FUNCTION "FRK_UnitRelease" : Void
{ S7_Optimized_Access := 'TRUE' }
VERSION : 0.1
VAR_INPUT
    Gate : DInt;
    Desired : DInt;
    Trusted : Bool;
    Core : "FRK_Core";
    Unit : "FRK_Unit";
    Status : "ST_ModuleStatus";
    Policy : Array[0..6] of "ST_ModePolicy";
    Access : "FRK_Access";
    Supported : Array[0..6] of Bool;
END_VAR
VAR_IN_OUT
    Report : "ST_ReleaseReport";
END_VAR
BEGIN
    #Report.Count := 0;
    #Report.Released := TRUE;
    IF #Gate <> 5 AND #Gate <> 4
        AND #Gate <> 7 AND #Gate <> 2
        AND #Gate <> 8
        AND NOT (#Unit.ConfigEnabled AND #Gate = 1)
        AND NOT (#Unit.ConfigSetsEnabled AND #Gate = 11)
        AND NOT (#Unit.ModelEnabled AND #Gate = 3) THEN
        "FRK_ReleaseReason"(Report := #Report, Description := WSTRING#'std.error.unsupportedHmiRequest', Reason := 2008, Path := STRING_TO_WSTRING(#Status.Name), Kind := 4);
        RETURN;
    END_IF;
    IF NOT #Trusted THEN
        IF #Access.CurrentLevel < #Access.Policy.Required[#Gate] THEN
            "FRK_ReleaseReason"(Report := #Report, Description := WSTRING#'std.release.insufficientAction', Reason := 2002, Path := STRING_TO_WSTRING(#Status.Name), Kind := 1);
        END_IF;
    END_IF;
    CASE #Gate OF
        3:
            IF #Core.Exec <> 0 OR #Unit.ModePending OR #Unit.Clearing OR NOT "FRK_DescendantsReady"(OwnerIndex := #Core.RegIndex) THEN
                "FRK_ReleaseReason"(Report := #Report, Description := WSTRING#'std.error.hmiRequestRejected', Reason := 2011, Path := STRING_TO_WSTRING(#Status.Name), Kind := 4);
            END_IF;
            IF #Unit.AlarmBlocking THEN
                "FRK_ReleaseReason"(Report := #Report, Description := WSTRING#'std.release.manualReset', Reason := 0, Path := STRING_TO_WSTRING(#Status.Name), Kind := 2);
            END_IF;
            IF NOT #Unit.Permit THEN
                "FRK_ReleaseReason"(Report := #Report, Description := #Unit.PermitDiag.Description, Reason := #Unit.PermitDiag.ReasonCode, Path := #Unit.PermitDiag.SourcePath, Kind := 3);
            END_IF;
        5:
            // Desired=0 is Start, Desired=1 is Stop. Generic action query is Stop.
            IF #Desired = 0 THEN
                IF #Unit.Mode = 1 OR #Unit.ModePending THEN
                    "FRK_ReleaseReason"(Report := #Report, Description := WSTRING#'std.error.unsupportedModeRequest', Reason := 2002, Path := STRING_TO_WSTRING(#Status.Name), Kind := 0);
                END_IF;
                IF #Core.Exec <> 0 OR #Unit.RunReq OR #Unit.Clearing OR #Unit.FaultLatched THEN
                    "FRK_ReleaseReason"(Report := #Report, Description := WSTRING#'std.error.hmiRequestRejected', Reason := 2011, Path := STRING_TO_WSTRING(#Status.Name), Kind := 4);
                END_IF;
                IF #Unit.AlarmBlocking THEN
                    "FRK_ReleaseReason"(Report := #Report, Description := WSTRING#'std.release.manualReset', Reason := 0, Path := STRING_TO_WSTRING(#Status.Name), Kind := 2);
                END_IF;
                IF #Unit.ConfigBlocked THEN
                    "FRK_ReleaseReason"(Report := #Report, Description := WSTRING#'std.release.configRestoreUnacknowledged', Reason := 2040, Path := STRING_TO_WSTRING(#Status.Name), Kind := 2);
                END_IF;
                IF NOT #Unit.Permit THEN
                    "FRK_ReleaseReason"(Report := #Report, Description := #Unit.PermitDiag.Description, Reason := #Unit.PermitDiag.ReasonCode, Path := #Unit.PermitDiag.SourcePath, Kind := 3);
                END_IF;
            END_IF;
        4:
            IF #Unit.ModePending THEN
                "FRK_ReleaseReason"(Report := #Report, Description := WSTRING#'std.release.modeChangeAlreadyPending', Reason := 2011, Path := STRING_TO_WSTRING(#Status.Name), Kind := 0);
            END_IF;
            IF #Core.Exec = 1 AND #Unit.Mode <> 1 THEN
                IF #Policy[#Unit.Mode].Shield = 2 THEN
                    "FRK_ReleaseReason"(Report := #Report, Description := WSTRING#'std.release.modeSwitchBlockedWhileRunning', Reason := 2002, Path := STRING_TO_WSTRING(#Status.Name), Kind := 0);
                END_IF;
            END_IF;
            IF #Desired <> -1 THEN
                IF #Desired < 0 OR #Desired >= 7 THEN
                    "FRK_ReleaseReason"(Report := #Report, Description := WSTRING#'std.error.unsupportedModeRequest', Reason := 2008, Path := STRING_TO_WSTRING(#Status.Name), Kind := 0);
                ELSIF NOT #Supported[#Desired] THEN
                    "FRK_ReleaseReason"(Report := #Report, Description := WSTRING#'std.error.unsupportedModeRequest', Reason := 2008, Path := STRING_TO_WSTRING(#Status.Name), Kind := 0);
                END_IF;
            END_IF;
        7:
            // The complete alarm model is separate; this gate owns the current latch.
            IF NOT #Unit.FaultLatched AND NOT #Unit.AlarmBlocking AND #Core.Exec = 0 AND NOT #Unit.Clearing AND NOT #Unit.ModePending AND NOT #Unit.FollowStart THEN
                IF "FRK_DescendantsReady"(OwnerIndex := #Core.RegIndex) THEN
                    "FRK_ReleaseReason"(Report := #Report, Description := WSTRING#'std.release.noBlockingAlarm', Reason := 2011, Path := STRING_TO_WSTRING(#Status.Name), Kind := 4);
                END_IF;
            END_IF;
        2:
            "FRK_ManualCommon"(Core := #Core, Unit := #Unit, Status := #Status, Report := #Report);
        ELSE
            RETURN;
    END_CASE;
END_FUNCTION

FUNCTION "FRK_ManualCommon" : Void
{ S7_Optimized_Access := 'TRUE' }
VERSION : 0.1
VAR_INPUT
    Core : "FRK_Core";
    Unit : "FRK_Unit";
    Status : "ST_ModuleStatus";
END_VAR
VAR_IN_OUT
    Report : "ST_ReleaseReport";
END_VAR
BEGIN
    IF #Unit.Mode <> 1 OR #Unit.ModePending THEN
        "FRK_ReleaseReason"(Report := #Report, Description := WSTRING#'std.release.manualModeRequired', Reason := 2002, Path := STRING_TO_WSTRING(#Status.Name), Kind := 0);
    END_IF;
    IF #Core.Exec <> 0 OR #Unit.Clearing OR #Unit.FaultLatched THEN
        "FRK_ReleaseReason"(Report := #Report, Description := WSTRING#'std.error.hmiRequestRejected', Reason := 2011, Path := STRING_TO_WSTRING(#Status.Name), Kind := 4);
    END_IF;
    IF #Unit.AlarmBlocking THEN
        "FRK_ReleaseReason"(Report := #Report, Description := WSTRING#'std.release.manualReset', Reason := 0, Path := STRING_TO_WSTRING(#Status.Name), Kind := 2);
    END_IF;
    IF NOT #Unit.Permit THEN
        "FRK_ReleaseReason"(Report := #Report, Description := #Unit.PermitDiag.Description, Reason := #Unit.PermitDiag.ReasonCode, Path := #Unit.PermitDiag.SourcePath, Kind := 3);
    END_IF;
END_FUNCTION

FUNCTION "FRK_ManualCondition" : Void
{ S7_Optimized_Access := 'TRUE' }
VERSION : 0.1
VAR_INPUT
    Slot : Int;
    Value : DInt;
    Ok : Bool;
    Diag : "ST_Diagnostic";
    Bypassable : Bool;
END_VAR
VAR_IN_OUT
    Conditions : Array[1..16] of "FRK_ManualConditionRow";
END_VAR
BEGIN
    IF #Slot < 1 OR #Slot > 16 THEN RETURN; END_IF;
    #Conditions[#Slot].Used := TRUE;
    #Conditions[#Slot].Value := #Value;
    #Conditions[#Slot].Ok := #Ok;
    #Conditions[#Slot].Diag := #Diag;
    #Conditions[#Slot].Bypassable := #Bypassable;
END_FUNCTION

FUNCTION "FRK_ManualApply" : Void
{ S7_Optimized_Access := 'TRUE' }
VERSION : 0.1
VAR_INPUT
    Request : "ST_HmiRequest";
    Status : "ST_ModuleStatus";
    Core : "FRK_Core";
    Commands : Array[1..12] of "ST_CommandInfo";
    Count : DInt;
    Conditions : Array[1..16] of "FRK_ManualConditionRow";
END_VAR
VAR_IN_OUT
    Report : "ST_ReleaseReport";
    Execute : Bool;
    Command : DInt;
    ManualOwned : Bool;
END_VAR
VAR_TEMP
    Index : Int;
    Supported : Bool;
    PreviousCount : Int;
END_VAR
BEGIN
    #Supported := FALSE;
    IF #Count >= 0 AND #Count <= 12 THEN
        FOR #Index := 1 TO DINT_TO_INT(#Count) DO
            IF #Commands[#Index].Value = #Request.IntValue AND #Commands[#Index].Style = 0 THEN #Supported := TRUE; END_IF;
        END_FOR;
    END_IF;
    IF NOT #Supported THEN
        "FRK_ReleaseReason"(Report := #Report, Description := WSTRING#'std.error.unsupportedHmiRequest', Reason := 2008, Path := STRING_TO_WSTRING(#Status.Name), Kind := 4);
    END_IF;
    IF #Core.Exec <> 0 OR #Execute OR #Core.ReleasePending THEN
        "FRK_ReleaseReason"(Report := #Report, Description := WSTRING#'std.error.hmiRequestRejected', Reason := 2011, Path := STRING_TO_WSTRING(#Status.Name), Kind := 4);
    END_IF;
    FOR #Index := 1 TO 16 DO
        IF #Conditions[#Index].Used AND NOT #Conditions[#Index].Ok THEN
            IF #Conditions[#Index].Value = 0 OR #Conditions[#Index].Value = #Request.IntValue THEN
                #PreviousCount := #Report.Count;
                "FRK_ReleaseReason"(Report := #Report, Description := #Conditions[#Index].Diag.Description, Reason := #Conditions[#Index].Diag.ReasonCode, Path := STRING_TO_WSTRING(#Status.Name), Kind := 3);
                IF #Report.Count > #PreviousCount THEN #Report.Reasons[#Report.Count].Bypassable := #Conditions[#Index].Bypassable; END_IF;
            END_IF;
        END_IF;
    END_FOR;
    IF #Request.Kind = 11 AND #Report.Released THEN
        #Command := #Request.IntValue;
        #Execute := TRUE;
        #ManualOwned := TRUE;
    END_IF;
END_FUNCTION

FUNCTION "FRK_ManualFinish" : Void
{ S7_Optimized_Access := 'TRUE' }
VERSION : 0.1
VAR_INPUT
    Core : "FRK_Core";
END_VAR
VAR_IN_OUT
    Execute : Bool;
    ManualOwned : Bool;
END_VAR
BEGIN
    IF #ManualOwned AND #Core.Exec <> 1 THEN
        #Execute := FALSE;
        #ManualOwned := FALSE;
    END_IF;
END_FUNCTION

FUNCTION "FRK_UnitCascade" : Void
{ S7_Optimized_Access := 'TRUE' }
VERSION : 0.1
VAR_INPUT
    ParentUnit : "FRK_Unit";
    Supported : Array[0..6] of Bool;
END_VAR
VAR_IN_OUT
    Core : "FRK_Core";
    Unit : "FRK_Unit";
    Status : "ST_ModuleStatus";
    Policy : Array[0..6] of "ST_ModePolicy";
    Access : "FRK_Access";
    AlarmLog : "FRK_AlarmLog";
END_VAR
VAR_TEMP
    Request : "ST_HmiRequest";
END_VAR
BEGIN
    IF NOT #ParentUnit.CascadePending THEN RETURN; END_IF;
    IF #ParentUnit.CascadeKind = 6 OR #ParentUnit.CascadeKind = 9 THEN
        #Unit.FollowStart := FALSE;
        #Request.Kind := #ParentUnit.CascadeKind;
        "FRK_UnitOperation"(Core := #Core, Unit := #Unit, Status := #Status, Policy := #Policy, Access := #Access, Supported := #Supported, Request := #Request, Response := "FRK_UnitScratch".Response, Trusted := TRUE);
        RETURN;
    END_IF;
    #Request.Kind := 3;
    #Request.IntValue := #ParentUnit.CascadeMode;
    "FRK_UnitOperation"(Core := #Core, Unit := #Unit, Status := #Status, Policy := #Policy, Access := #Access, Supported := #Supported, Request := #Request, Response := "FRK_UnitScratch".Response, Trusted := TRUE);
    IF NOT "FRK_UnitScratch".Response.Accepted THEN
        #Unit.FollowStart := FALSE;
        #Request.Kind := 6;
        "FRK_UnitOperation"(Core := #Core, Unit := #Unit, Status := #Status, Policy := #Policy, Access := #Access, Supported := #Supported, Request := #Request, Response := "FRK_UnitScratch".Response, Trusted := TRUE);
        // Core names this event but has no assigned E_Reason ordinal yet.
        "FRK_AlarmMessage"(AlarmLog := #AlarmLog, Reason := 2008, Description := WSTRING#'std.event.childModeUnsupported', SourcePath := STRING_TO_WSTRING(#Status.Name));
    ELSE
        #Unit.FollowStart := #ParentUnit.CascadeKind = 5;
    END_IF;
END_FUNCTION

FUNCTION "FRK_UnitFollow" : Void
{ S7_Optimized_Access := 'TRUE' }
VERSION : 0.1
VAR_INPUT
    Supported : Array[0..6] of Bool;
END_VAR
VAR_IN_OUT
    Core : "FRK_Core";
    Unit : "FRK_Unit";
    Status : "ST_ModuleStatus";
    Policy : Array[0..6] of "ST_ModePolicy";
    Access : "FRK_Access";
END_VAR
VAR_TEMP
    Request : "ST_HmiRequest";
END_VAR
BEGIN
    IF #Unit.FollowStart AND NOT #Unit.ModePending AND NOT #Unit.Clearing THEN
        #Unit.FollowStart := FALSE;
        #Request.Kind := 5;
        "FRK_UnitOperation"(Core := #Core, Unit := #Unit, Status := #Status, Policy := #Policy, Access := #Access, Supported := #Supported, Request := #Request, Response := "FRK_UnitScratch".Response, Trusted := TRUE);
    END_IF;
END_FUNCTION

// Core 6.11: one authoritative decision slot per registered root.
FUNCTION "FRK_DecisionRoot" : Int
{ S7_Optimized_Access := 'TRUE' }
VERSION : 0.1
VAR_INPUT Owner : DInt; Create : Bool; END_VAR
VAR_TEMP RootIndex : DInt; Depth : DInt; Slot : Int; END_VAR
BEGIN
    #FRK_DecisionRoot := 0;
    IF "FRK_Registry".Fault OR "FRK_Registry".Count < 1 OR "FRK_Registry".Count > 4 THEN RETURN; END_IF;
    #RootIndex := #Owner;
    FOR #Depth := 1 TO 4 DO
        IF #RootIndex < 1 OR #RootIndex > "FRK_Registry".Count THEN RETURN; END_IF;
        IF NOT "FRK_Registry".Rows[#RootIndex].Valid THEN RETURN; END_IF;
        IF "FRK_Registry".Rows[#RootIndex].Parent = 0 THEN EXIT; END_IF;
        #RootIndex := "FRK_Registry".Rows[#RootIndex].Parent;
    END_FOR;
    IF "FRK_Registry".Rows[#RootIndex].Parent <> 0 THEN RETURN; END_IF;
    FOR #Slot := 1 TO 1 DO
        IF "FRK_Decisions".Slots[#Slot].RootIndex = #RootIndex THEN
            #FRK_DecisionRoot := #Slot;
            RETURN;
        END_IF;
    END_FOR;
    IF NOT #Create THEN RETURN; END_IF;
    FOR #Slot := 1 TO 1 DO
        IF "FRK_Decisions".Slots[#Slot].RootIndex = 0 THEN
            "FRK_Decisions".Slots[#Slot].RootIndex := #RootIndex;
            #FRK_DecisionRoot := #Slot;
            RETURN;
        END_IF;
    END_FOR;
END_FUNCTION

FUNCTION "FRK_DecisionAudit" : Void
{ S7_Optimized_Access := 'TRUE' }
VERSION : 0.1
VAR_INPUT Key : WString; SourcePath : WString; Option : Int; END_VAR
VAR_IN_OUT AlarmLog : "FRK_AlarmLog"; END_VAR
VAR_TEMP Diag : "ST_Diagnostic"; Slot : Int; Gone : Bool; END_VAR
BEGIN
    #Diag := "FRK_UnitScratch".EmptyDiagnostic;
    #Diag.Description := #Key;
    IF #Option <> 0 THEN
        #Diag.Description := CONCAT(IN1 := #Diag.Description, IN2 := WSTRING#' option=');
        #Diag.Description := CONCAT(IN1 := #Diag.Description, IN2 := STRING_TO_WSTRING(INT_TO_STRING(#Option)));
    END_IF;
    #Diag.SourcePath := #SourcePath;
    #Diag.Severity := 0;
    #Diag.Category := 0;
    #Slot := "FRK_AlarmRaise"(AlarmLog := #AlarmLog, Diag := #Diag, ResetClass := 0);
    IF #Slot > 0 THEN #Gone := "FRK_AlarmGone"(AlarmLog := #AlarmLog, Slot := #Slot); END_IF;
END_FUNCTION

FUNCTION "FRK_DecisionClear" : Void
{ S7_Optimized_Access := 'TRUE' }
VERSION : 0.1
VAR_IN_OUT Slot : "FRK_DecisionSlot"; END_VAR
VAR_TEMP Index : Int; END_VAR
BEGIN
    #Slot.Request.Prompt := WSTRING#'';
    #Slot.Request.SourcePath := WSTRING#'';
    #Slot.Request.Default := 0;
    #Slot.Request.Timeout := T#0ms;
    FOR #Index := 1 TO 6 DO #Slot.Request.Options[#Index] := ''; END_FOR;
    #Slot.Answer := 0;
    #Slot.Owner := 0;
    #Slot.OverlapLogged := FALSE;
    #Slot.ResolutionLogged := FALSE;
END_FUNCTION

FUNCTION "FRK_DecisionAsk" : Bool
{ S7_Optimized_Access := 'TRUE' }
VERSION : 0.1
VAR_INPUT Owner : DInt; OwnerPath : WString; Request : "ST_DecisionRequest"; END_VAR
VAR_IN_OUT AlarmLog : "FRK_AlarmLog"; END_VAR
VAR_TEMP Candidate : "ST_DecisionRequest"; Slot : Int; Index : Int; SameRequest : Bool; HasOption : Bool; END_VAR
BEGIN
    #FRK_DecisionAsk := FALSE;
    #Slot := "FRK_DecisionRoot"(Owner := #Owner, Create := TRUE);
    IF #Slot = 0 THEN RETURN; END_IF;
    #Candidate := #Request;
    IF #Candidate.SourcePath = WSTRING#'' THEN
        #Candidate.SourcePath := #OwnerPath;
    END_IF;
    IF "FRK_Decisions".Slots[#Slot].Request.Prompt <> WSTRING#'' THEN
        #SameRequest := "FRK_Decisions".Slots[#Slot].Owner = #Owner
            AND "FRK_Decisions".Slots[#Slot].Request.Prompt = #Candidate.Prompt
            AND "FRK_Decisions".Slots[#Slot].Request.SourcePath = #Candidate.SourcePath
            AND "FRK_Decisions".Slots[#Slot].Request.Default = #Candidate.Default
            AND "FRK_Decisions".Slots[#Slot].Request.Timeout = #Candidate.Timeout;
        FOR #Index := 1 TO 6 DO
            #SameRequest := #SameRequest AND "FRK_Decisions".Slots[#Slot].Request.Options[#Index] = #Candidate.Options[#Index];
        END_FOR;
        IF #SameRequest THEN #FRK_DecisionAsk := TRUE; RETURN; END_IF;
        IF NOT "FRK_Decisions".Slots[#Slot].OverlapLogged THEN
            "FRK_DecisionAudit"(AlarmLog := #AlarmLog, Key := WSTRING#'std.audit.decisionOverlapRejected', SourcePath := #Candidate.SourcePath, Option := 0);
            "FRK_Decisions".Slots[#Slot].OverlapLogged := TRUE;
        END_IF;
        RETURN;
    END_IF;
    #HasOption := FALSE;
    FOR #Index := 1 TO 6 DO #HasOption := #HasOption OR #Candidate.Options[#Index] <> ''; END_FOR;
    IF #Candidate.Prompt = WSTRING#'' OR #Candidate.Timeout < T#0ms OR NOT #HasOption
        OR #Candidate.SourcePath <> #OwnerPath OR #OwnerPath = WSTRING#'' THEN
        "FRK_DecisionAudit"(AlarmLog := #AlarmLog, Key := WSTRING#'std.audit.decisionInvalidRejected', SourcePath := #Candidate.SourcePath, Option := #Candidate.Default);
        RETURN;
    END_IF;
    IF #Candidate.Timeout > T#0ms OR #Candidate.Default <> 0 THEN
        IF #Candidate.Default < 1 OR #Candidate.Default > 6 THEN
            "FRK_DecisionAudit"(AlarmLog := #AlarmLog, Key := WSTRING#'std.audit.decisionInvalidRejected', SourcePath := #Candidate.SourcePath, Option := #Candidate.Default);
            RETURN;
        END_IF;
        IF #Candidate.Options[#Candidate.Default] = '' THEN
            "FRK_DecisionAudit"(AlarmLog := #AlarmLog, Key := WSTRING#'std.audit.decisionInvalidRejected', SourcePath := #Candidate.SourcePath, Option := #Candidate.Default);
            RETURN;
        END_IF;
    END_IF;
    "FRK_Decisions".Slots[#Slot].Request := #Candidate;
    "FRK_Decisions".Slots[#Slot].Owner := #Owner;
    "FRK_Decisions".Slots[#Slot].AskedAt := "FRK_Clock".NowMs;
    "FRK_Decisions".Slots[#Slot].Answer := 0;
    "FRK_Decisions".Slots[#Slot].ResolutionLogged := FALSE;
    "FRK_Decisions".Slots[#Slot].OverlapLogged := FALSE;
    "FRK_DecisionAudit"(AlarmLog := #AlarmLog, Key := WSTRING#'std.audit.decisionRequested', SourcePath := #Candidate.SourcePath, Option := 0);
    #FRK_DecisionAsk := TRUE;
END_FUNCTION

FUNCTION "FRK_DecisionSubmit" : Bool
{ S7_Optimized_Access := 'TRUE' }
VERSION : 0.1
VAR_INPUT Owner : DInt; OwnerPath : WString; Option : DInt; Busy : Bool; Permit : Bool; END_VAR
VAR_IN_OUT Report : "ST_ReleaseReport"; END_VAR
VAR_TEMP Slot : Int; SourcePath : WString[255]; END_VAR
BEGIN
    #FRK_DecisionSubmit := FALSE;
    #Slot := "FRK_DecisionRoot"(Owner := #Owner, Create := FALSE);
    #SourcePath := #OwnerPath;
    IF NOT #Busy OR #Slot = 0 THEN
        "FRK_ReleaseReason"(Report := #Report, Description := WSTRING#'std.release.noActiveDecision', Reason := 0, Path := #SourcePath, Kind := 4);
        RETURN;
    END_IF;
    IF "FRK_Decisions".Slots[#Slot].RootIndex <> #Owner THEN
        "FRK_ReleaseReason"(Report := #Report, Description := WSTRING#'std.release.noActiveDecision', Reason := 0, Path := #SourcePath, Kind := 4);
        RETURN;
    END_IF;
    IF "FRK_Decisions".Slots[#Slot].Request.Prompt = WSTRING#'' OR "FRK_Decisions".Slots[#Slot].Answer <> 0 THEN
        "FRK_ReleaseReason"(Report := #Report, Description := WSTRING#'std.release.noActiveDecision', Reason := 0, Path := #SourcePath, Kind := 4);
        RETURN;
    END_IF;
    IF #Option < 1 OR #Option > 6 THEN
        "FRK_ReleaseReason"(Report := #Report, Description := WSTRING#'std.release.invalidDecisionOption', Reason := 2008, Path := #SourcePath, Kind := 4);
        RETURN;
    END_IF;
    IF "FRK_Decisions".Slots[#Slot].Request.Options[#Option] = '' THEN
        "FRK_ReleaseReason"(Report := #Report, Description := WSTRING#'std.release.invalidDecisionOption', Reason := 2008, Path := #SourcePath, Kind := 4);
        RETURN;
    END_IF;
    IF NOT #Permit THEN
        "FRK_ReleaseReason"(Report := #Report, Description := WSTRING#'std.release.decisionInterlock', Reason := 2002, Path := #SourcePath, Kind := 3);
        RETURN;
    END_IF;
    IF NOT #Report.Released THEN RETURN; END_IF;
    "FRK_Decisions".Slots[#Slot].Answer := DINT_TO_INT(#Option);
    #FRK_DecisionSubmit := TRUE;
END_FUNCTION

FUNCTION "FRK_DecisionCyclic" : Void
{ S7_Optimized_Access := 'TRUE' }
VERSION : 0.1
VAR_INPUT Owner : DInt; Busy : Bool; Reset : Bool; END_VAR
VAR_IN_OUT AlarmLog : "FRK_AlarmLog"; END_VAR
VAR_TEMP Slot : Int; Elapsed : UDInt; END_VAR
BEGIN
    IF #Owner < 1 OR #Owner > "FRK_Registry".Count THEN RETURN; END_IF;
    // Only the root resolves/withdraws its slot; an idle nested Unit cannot
    // cancel a root's running decision.
    IF "FRK_Registry".Rows[#Owner].Parent <> 0 THEN RETURN; END_IF;
    #Slot := "FRK_DecisionRoot"(Owner := #Owner, Create := FALSE);
    IF #Slot = 0 THEN RETURN; END_IF;
    IF "FRK_Decisions".Slots[#Slot].Request.Prompt = WSTRING#'' THEN RETURN; END_IF;
    IF #Reset OR NOT #Busy THEN
        "FRK_DecisionAudit"(AlarmLog := #AlarmLog, Key := WSTRING#'std.audit.decisionWithdrawn', SourcePath := "FRK_Decisions".Slots[#Slot].Request.SourcePath, Option := 0);
        "FRK_DecisionClear"(Slot := "FRK_Decisions".Slots[#Slot]);
        RETURN;
    END_IF;
    IF "FRK_Decisions".Slots[#Slot].Answer <> 0 THEN
        IF NOT "FRK_Decisions".Slots[#Slot].ResolutionLogged THEN
            "FRK_DecisionAudit"(AlarmLog := #AlarmLog, Key := WSTRING#'std.audit.decisionOperatorResolved', SourcePath := "FRK_Decisions".Slots[#Slot].Request.SourcePath, Option := "FRK_Decisions".Slots[#Slot].Answer);
            "FRK_Decisions".Slots[#Slot].ResolutionLogged := TRUE;
        END_IF;
        RETURN;
    END_IF;
    IF "FRK_Decisions".Slots[#Slot].Request.Timeout <= T#0ms THEN RETURN; END_IF;
    #Elapsed := "FRK_Clock".NowMs - "FRK_Decisions".Slots[#Slot].AskedAt;
    IF #Elapsed >= DINT_TO_UDINT(TIME_TO_DINT("FRK_Decisions".Slots[#Slot].Request.Timeout)) THEN
        "FRK_Decisions".Slots[#Slot].Answer := "FRK_Decisions".Slots[#Slot].Request.Default;
        "FRK_DecisionAudit"(AlarmLog := #AlarmLog, Key := WSTRING#'std.audit.decisionTimeoutResolved', SourcePath := "FRK_Decisions".Slots[#Slot].Request.SourcePath, Option := "FRK_Decisions".Slots[#Slot].Answer);
        "FRK_Decisions".Slots[#Slot].ResolutionLogged := TRUE;
    END_IF;
END_FUNCTION

FUNCTION "FRK_DecisionTake" : Int
{ S7_Optimized_Access := 'TRUE' }
VERSION : 0.1
VAR_INPUT Owner : DInt; END_VAR
VAR_IN_OUT AlarmLog : "FRK_AlarmLog"; END_VAR
VAR_TEMP Slot : Int; END_VAR
BEGIN
    #FRK_DecisionTake := 0;
    #Slot := "FRK_DecisionRoot"(Owner := #Owner, Create := FALSE);
    IF #Slot = 0 THEN RETURN; END_IF;
    IF "FRK_Decisions".Slots[#Slot].Owner <> #Owner THEN RETURN; END_IF;
    IF "FRK_Decisions".Slots[#Slot].Answer = 0 THEN RETURN; END_IF;
    #FRK_DecisionTake := "FRK_Decisions".Slots[#Slot].Answer;
    IF NOT "FRK_Decisions".Slots[#Slot].ResolutionLogged THEN
        "FRK_DecisionAudit"(AlarmLog := #AlarmLog, Key := WSTRING#'std.audit.decisionOperatorResolved', SourcePath := "FRK_Decisions".Slots[#Slot].Request.SourcePath, Option := #FRK_DecisionTake);
    END_IF;
    "FRK_DecisionClear"(Slot := "FRK_Decisions".Slots[#Slot]);
END_FUNCTION

FUNCTION "FRK_DecisionPublish" : Void
{ S7_Optimized_Access := 'TRUE' }
VERSION : 0.1
VAR_INPUT Owner : DInt; END_VAR
VAR_IN_OUT Decision : "ST_DecisionRequest"; DecisionAnswer : Int; END_VAR
VAR_TEMP Slot : Int; END_VAR
BEGIN
    #Slot := "FRK_DecisionRoot"(Owner := #Owner, Create := FALSE);
    #Decision := "FRK_Decisions".EmptyRequest;
    #DecisionAnswer := 0;
    IF #Slot = 0 THEN RETURN; END_IF;
    IF "FRK_Decisions".Slots[#Slot].RootIndex <> #Owner THEN RETURN; END_IF;
    #Decision := "FRK_Decisions".Slots[#Slot].Request;
    #DecisionAnswer := "FRK_Decisions".Slots[#Slot].Answer;
END_FUNCTION
